{attribute 'qualified_only'}
{attribute 'strict'}
TYPE E_CIP_Return :
(
	eNone := 0,
	eDrain,
	eT91_Sanitation,
	eT92_Detergent,
	eT93_R_Water,
	eT94_Water
);
END_TYPE

(* stored: Version 1.1.0.1, ProductVersion 3.1.4024.12
   DUT E_CIP_Return: Id {86496414-0861-4ef3-a003-80b87181b00c} *)
